// TwinCAT 3 PLC project CX7080_Robot_Controller
// ProgramVersion: 3.1.4024.0
// libraries:
//   Tc2_ModbusRTU, * (Beckhoff Automation GmbH)
//   Tc2_Standard, * (Beckhoff Automation GmbH)
//   Tc2_System, * (Beckhoff Automation GmbH)
//   Tc2_Utilities, * (Beckhoff Automation GmbH)
//   Tc3_Module, * (Beckhoff Automation GmbH)
// project tree:
//   DUTs/ eMbCycleState.TcDUT, eMbDiag.TcDUT, ST_HW_DI.TcDUT, ST_HW_DO.TcDUT, ST_MB_ReadRegs.TcDUT, ST_MB_WriteRegs.TcDUT, state_enum.TcDUT
//   GVLs/ GVL.TcGVL
//   / PlcTask.TcTTO
//   POUs/Comms/ FB_i_Watchdog.TcPOU, FB_ModbusComm.TcPOU, FB_Toggle_ReadWrite.TcPOU
//   POUs/ FB_Startup.TcPOU, I_JointJog.TcIO, MAIN.TcPOU, TESTING.TcPOU
//   POUs/Misc/ FB_System_Time.TcPOU
//   POUs/Motion/ FB_AutoSequence.TcPOU, FB_Jog_Joint.TcPOU, FB_Servo.TcPOU
//   POUs/Utilities/ FB_ElectromagnetActivate.TcPOU
// real-time tasks:
//   TASK PlcTask: cycle T#10ms, priority 20, ADS port 350
//   TASK PlcTask1: cycle T#10ms, priority 21, ADS port 351
//   TASK PlcTask2: cycle T#10ms, priority 22, ADS port 352
// I/O:
//   DEVICE Device 3 (CX7000), AmsNetId 5.140.122.236.4.1
//     Term 1 (CX7028) [CX7028-0000-0121]
//       modules: Module 1 (DIO_2x), Module 2 (Empty Module), Module 3 (DIO_2x), Module 4 (Empty Module), Module 5 (DI_2x), Module 6 (Empty Module), Module 7 (DI_2x), Module 8 (Empty Module)
//   DEVICE Device 1 (EtherCAT), AmsNetId 5.140.122.236.2.1
//     Term 1 (EK1200) [EK1200-7000 EtherCAT Power supply (1,5A E-Bus)]
//       Term 2 (EL1008) [EL1008 8Ch. Dig. Input 24V, 3ms]
//       Term 3 (EL1008) [EL1008 8Ch. Dig. Input 24V, 3ms]
//       Term 4 (EL2008) [EL2008 8Ch. Dig. Output 24V, 0.5A]
//       Term 5 (EL2008) [EL2008 8Ch. Dig. Output 24V, 0.5A]
//   DEVICE Device 7 (COM Port)
// variable links:
//   CX7080_Robot_Controller Instance <-> Device 1 (EtherCAT)/Term 1 (EK1200)/Term 2 (EL1008)
//     PlcTask Inputs/GVL.PB_EE_Grip <-> Channel 6/Input
//     PlcTask Inputs/GVL.PB_EE_Ungrip <-> Channel 8/Input
//     PlcTask Inputs/GVL.PB_J1_CCW <-> Channel 3/Input
//     PlcTask Inputs/GVL.PB_J2_CCW <-> Channel 5/Input
//     PlcTask Inputs/GVL.PB_J3_CCW <-> Channel 2/Input
//     PlcTask Inputs/GVL.PB_J1_CW <-> Channel 1/Input
//     PlcTask Inputs/GVL.PB_J2_CW <-> Channel 7/Input
//     PlcTask Inputs/GVL.PB_J3_CW <-> Channel 4/Input
//   CX7080_Robot_Controller Instance <-> Device 1 (EtherCAT)/Term 1 (EK1200)/Term 3 (EL1008)
//     PlcTask Inputs/GVL.PB_EMG_STOP <-> Channel 1/PB_EMG_STOP
//     PlcTask Inputs/GVL.PB_Record_Pos <-> Channel 3/PB_RECORD_POS
//     PlcTask Inputs/GVL.PB_Reset <-> Channel 2/PB_RESET
//     PlcTask Inputs/GVL.PB_Start_Pause <-> Channel 5/PB_START_PAUSE
//     PlcTask Inputs/GVL.SW_Jog_Auto <-> Channel 6/SW_JOG_AUTO
//     PlcTask Inputs/GVL.SW_Join_Cart <-> Channel 8/SW_JOINT_CART
//     PlcTask Inputs/GVL.SW_Slow_Fast <-> Channel 4/SW_SLOW_FAST
//   CX7080_Robot_Controller Instance <-> Device 1 (EtherCAT)/Term 1 (EK1200)/Term 4 (EL2008)
//     PlcTask Outputs/GVL.LED_EE_Grip <-> Channel 6/Output
//     PlcTask Outputs/GVL.LED_EE_Ungrip <-> Channel 8/Output
//     PlcTask Outputs/GVL.LED_J1_CCW <-> Channel 3/Output
//     PlcTask Outputs/GVL.LED_J2_CCW <-> Channel 5/Output
//     PlcTask Outputs/GVL.LED_J3_CCW <-> Channel 2/Output
//     PlcTask Outputs/GVL.LED_J1_CW <-> Channel 1/Output
//     PlcTask Outputs/GVL.LED_J2_CW <-> Channel 7/Output
//     PlcTask Outputs/GVL.LED_J3_CW <-> Channel 4/Output
//   CX7080_Robot_Controller Instance <-> Device 1 (EtherCAT)/Term 1 (EK1200)/Term 5 (EL2008)
//     PlcTask Outputs/GVL.LED_Comm_Fault <-> Channel 6/Output
//     PlcTask Outputs/GVL.LED_EMG_STOP <-> Channel 1/Output
//     PlcTask Outputs/GVL.LED_Record_Pos <-> Channel 3/Output
//     PlcTask Outputs/GVL.LED_Reset <-> Channel 2/Output
//     PlcTask Outputs/GVL.LED_Start_Pause <-> Channel 5/Output
//     PlcTask Outputs/GVL.LED_Warning <-> Channel 7/Output
//   CX7080_Robot_Controller Instance <-> Device 7 (COM Port)
//     PlcTask Inputs/MAIN.fb_ModbusComm.MB_Master.InData @bit {16..520 step 8} <-> Inputs/Data{1..64}  (64 links)
//     PlcTask Inputs/MAIN.fb_ModbusComm.MB_Master.InData <-> Inputs/Status
//     PlcTask Outputs/MAIN.fb_ModbusComm.MB_Master.OutData <-> Outputs/Ctrl
//     PlcTask Outputs/MAIN.fb_ModbusComm.MB_Master.OutData @bit {16..520 step 8} <-> Outputs/Data{1..64}  (64 links)

CONFIGURATION CX7080_Robot_Controller
    RESOURCE PLC ON TwinCAT3
        TASK PlcTask(INTERVAL := T#10ms, PRIORITY := 22);
        PROGRAM MAIN WITH PlcTask : MAIN;
    END_RESOURCE
END_CONFIGURATION

// ---- DUTs/eMbCycleState.TcDUT
{attribute 'namespace' := 'MyLib.Modbus'}
TYPE eMbCycleState :
(
    eMbState_Init,
    eMbState_Read,
    eMbState_Write,
    eMbState_Error
);
END_TYPE

// ---- DUTs/eMbDiag.TcDUT
TYPE eMbDiag :
(
    eMbDiag_Ok := 0,
    eMbDiag_Timeout := 1,
    eMbDiag_InvalidBusy := 2
);
END_TYPE

// ---- DUTs/ST_HW_DI.TcDUT
TYPE ST_HW_DI :
STRUCT
END_STRUCT
END_TYPE

// ---- DUTs/ST_HW_DO.TcDUT
TYPE ST_HW_DO :
STRUCT
END_STRUCT
END_TYPE

// ---- DUTs/ST_MB_ReadRegs.TcDUT
TYPE ST_MB_ReadRegs :
STRUCT
END_STRUCT
END_TYPE

// ---- DUTs/ST_MB_WriteRegs.TcDUT
TYPE ST_MB_WriteRegs :
STRUCT
END_STRUCT
END_TYPE

// ---- DUTs/state_enum.TcDUT
{attribute 'qualified_only'}
{attribute 'strict'}
TYPE state_enum :
(
	startup_mode,
	jog_joint_mode,
	jog_cartesian_mode,
	auto_mode,
	emg_stop_mode,
	comm_fault_mode,
	manual_mode
);
END_TYPE

// ---- GVLs/GVL.TcGVL
{attribute 'qualified_only'}
VAR_GLOBAL
	// Internal system parameters
	system_state : state_enum := state_enum.startup_mode; // Used to keep track of system state machine. Initialized in startup_mode.
	modbus_comm_fault : BOOL := FALSE;
	J1_Home_Pos : INT := 135; // Degrees
	J2_Home_Pos : INT := 135; // Degrees
	J3_Home_Pos : INT := 135; // Degrees
	LowSpeedSetting : REAL := 5; // [deg/s]
	HighSpeedSetting : REAL := 20; // [deg/s]
	
	BaseAngleMin : INT := 0;
	BaseAngleMax : INT := 180;
	ShoulderAngleMin : INT := 20;
	ShoulderAngleMax : INT := 120;
	ElbowAngleMin : INT := 0;
	ElbowAngleMax : INT := 180;
	
	// Inputs
	input1 AT %I* : BOOL;
	output1 AT %Q* : BOOL;
	PB_J1_CW AT %I* : BOOL;
	PB_J1_CCW AT %I*: BOOL;
	PB_J2_CW AT %I* : BOOL;
	PB_J2_CCW AT %I* : BOOL;
	PB_J3_CW AT %I* : BOOL;
	PB_J3_CCW AT %I* : BOOL;
	PB_EE_Grip AT %I* : BOOL;
	PB_EE_Ungrip AT %I* : BOOL;
	PB_EMG_STOP AT %I* : BOOL;
	PB_Reset AT %I* : BOOL;
	PB_Record_Pos AT %I* : BOOL;
	PB_Record_Delay AT %I* : BOOL;
	PB_Start_Pause AT %I* : BOOL;
	SW_Slow_Fast AT %I* : BOOL;
	SW_Join_Cart AT %I* : BOOL;
	SW_Jog_Auto AT %I* : BOOL;
	
	// Outputs
	LED_J1_CW AT %Q* : BOOL;
	LED_J1_CCW AT %Q*: BOOL;
	LED_J2_CW AT %Q* : BOOL;
	LED_J2_CCW AT %Q* : BOOL;
	LED_J3_CW AT %Q* : BOOL;
	LED_J3_CCW AT %Q* : BOOL;
	LED_EE_Grip AT %Q* : BOOL;
	LED_EE_Ungrip AT %Q* : BOOL;
	LED_EMG_STOP AT %Q* : BOOL;
	LED_Reset AT %Q* : BOOL;
	LED_Record_Pos AT %Q* : BOOL;
	LED_Record_Delay AT %Q* : BOOL;
	LED_Start_Pause AT %Q* : BOOL;
	LED_Comm_Fault AT %Q* : BOOL;
	LED_Warning AT %Q* : BOOL;
	
	// Modbus registers
	MB_Write_J1 : INT;
	MB_Write_J2 : INT;
	MB_Write_J3 : INT;
	MB_Write_Gripper : INT;
	MB_Write_Watchdog : INT;
	MB_Write_Blank1 : INT;
	MB_Write_Blank2 : INT;
	MB_Write_Blank3 : INT;
	MB_Write_Blank4 : INT;
	MB_Write_Blank5 : INT;
	MB_Read_Watchdog : INT;
	MB_Read_Blank2 : INT;
	MB_Read_Blank3 : INT;
	MB_Read_Blank4 : INT;
	MB_Read_Blank5 : INT;
	MB_Read_Blank6 : INT;
	MB_Read_Blank7 : INT;
	MB_Read_Blank8 : INT;
	MB_Read_Blank9 : INT;
	MB_Read_Blank10 : INT;
	
END_VAR

// ---- POUs/I_JointJog.TcIO
INTERFACE I_JointJog


(*
Hva er poenget med å bruke interface?
Det gjør separation of concerns enklere.
En funksjonsblokk trenger ikke å vite hvordan ting er implementert i (en annen funksjonsblokk?), men trenger
bare å kjenne til interface.
Dette gjør det enklere å drive med TDD (test driven development), da funksjonsblokker har mindre avhengigheter.


*)

METHOD Ramp : LREAL
VAR_INPUT
END_VAR
END_METHOD

END_INTERFACE

// ---- POUs/MAIN.TcPOU
PROGRAM MAIN
VAR
	fb_Startup : FB_Startup;
	fb_ModbusComm: FB_ModbusComm;
	fb_System_Time : FB_System_Time;
	fb_Jog_Joint : FB_Jog_Joint;
	fb_ElectromagnetActivate : FB_ElectromagnetActivate;
END_VAR


(*
GJENSTÅENDE ARBEID:
1) Implementer auto sekvens FB
2) 
*)


GVL.LED_J1_CW := GVL.PB_J1_CW;
GVL.LED_J2_CW := GVL.PB_J2_CW;
GVL.LED_J3_CW := GVL.PB_J3_CW;
GVL.LED_J1_CCW := GVL.PB_J1_CCW;
GVL.LED_J2_CCW := GVL.PB_J2_CCW;
GVL.LED_J3_CCW := GVL.PB_J3_CCW;
GVL.LED_EE_Grip := GVL.PB_EE_Grip;
GVL.LED_EE_Ungrip := GVL.PB_EE_Ungrip;
GVL.LED_EMG_STOP := NOT GVL.PB_EMG_STOP;
GVL.LED_Start_Pause := GVL.PB_Start_Pause;
GVL.LED_Reset := GVL.LED_Reset;
GVL.LED_Warning := TRUE;
GVL.LED_Reset := GVL.PB_Reset;
GVL.LED_Start_Pause := GVL.PB_Start_Pause;
GVL.LED_Record_Pos := GVL.PB_Record_Pos;


// Code which must run every PLC cycle.
fb_System_Time(); // Run FB to calculate Delta_Time


(* COMMENTING OUT FOR TESTING PURPOSES
IF NOT GVL.PB_EMG_STOP AND NOT (gvl.system_state = state_enum.startup_mode) THEN
	GVL.system_state := state_enum.emg_stop_mode;
ELSIF GVL.LED_Comm_Fault AND NOT (gvl.system_state = state_enum.startup_mode)  THEN
	GVL.system_state := state_enum.comm_fault_mode;
END_IF
*)


CASE gvl.system_state OF
state_enum.startup_mode:
	fb_Startup();
state_enum.jog_joint_mode:
	fb_Jog_Joint(
	lr_DeltaTime:= fb_ModbusComm.lreal_CycleTime, 
	lr_SlowModeVelocitySetting:= 1, 
	lr_FastModeVelovitySetting:= 10, 
	i_Base_LowLimit:= 0, 
	i_Base_HighLimit:= 180, 
	i_Shoulder_LowLimit:= 0, 
	i_Shoulder_HighLimit:= 180, 
	i_Elbow_LowLimit:= 0, 
	i_Elbow_HighLimit:= 180, 
	b_Enable_Servos:= TRUE, 
	SW_Fast_Mode:= GVL.SW_Slow_Fast, 
	PB_Base_Pos:= GVL.PB_J1_CCW, 
	PB_Base_Neg:= GVL.PB_J1_CW, 
	PB_Shoulder_Pos:= GVL.PB_J2_CCW, 
	PB_Shoulder_Neg:= GVL.PB_J2_CW, 
	PB_Elbow_Pos:= GVL.PB_J3_CCW, 
	PB_Elbow_Neg:= GVL.PB_J3_CW, 
	i_Set_Base=>, 
	i_Set_Shoulder=>, 
	i_Set_Elbow=>);
	
	fb_ElectromagnetActivate(
	b_activate := GVL.PB_EE_Grip,
	b_deactivate := GVL.PB_EE_Ungrip,
	b_CMD_Magnet =>);
	
state_enum.jog_cartesian_mode:
state_enum.manual_mode:
state_enum.emg_stop_mode:
state_enum.comm_fault_mode:
state_enum.auto_mode:
END_CASE

//fb_ModbusComm();
fb_ModbusComm(
	i_MBO_BaseAngle:= fb_Jog_Joint.i_Set_Base, 
	i_MBO_ShoulderAngle:= fb_Jog_Joint.i_Set_Shoulder, 
	i_MBO_ElbowAngle:= fb_Jog_Joint.i_Set_Elbow, 
	i_MBO_EndEffectorValue:= BOOL_TO_INT(fb_ElectromagnetActivate.b_CMD_Magnet), 
	b_MBO_EmergencyStop:= , 
	lreal_CycleTime := fb_System_Time.Delta_Time,
	iLastWrittenBaseAngle=> , 
	iLastWrittenShoulderAngle=> , 
	iLastWrittenElbowAngle=> , 
	b_MBI_LocalControl=> , 
	b_MBI_LocalEmergencyStopActive=> , 
	b_MBWatchdogTimeout=> GVL.LED_Comm_Fault, 
	i_MBI_LocalBaseAngle=> , 
	i_MBI_LocalShoulderAngle=> , 
	i_MBI_LocalElbowAngle=> , 
	i_MBI_LocalValueEndEffector=> );

END_PROGRAM

// ---- POUs/FB_Startup.TcPOU
FUNCTION_BLOCK FB_Startup
VAR_INPUT
END_VAR
VAR_OUTPUT
END_VAR
VAR
	timer1 : TON;
	timer2 : TON;
	timer3 : TON;
	timer4 : TON;
	timer5 : TON;
	timer6 : TON;
	timer7 : TON;
	EMG_STOP_RELEASED : BOOL;
END_VAR

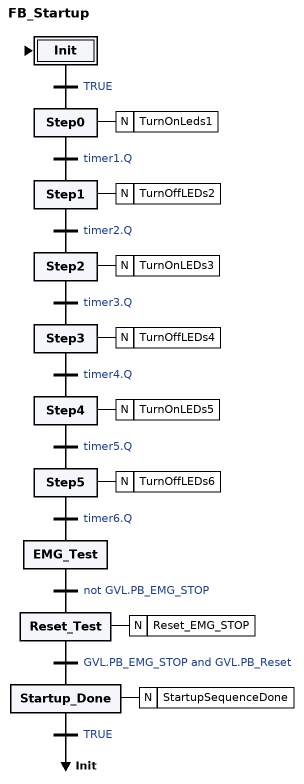
INITIAL_STEP Init:
END_STEP
TRANSITION FROM Init TO Step0
    := TRUE;
END_TRANSITION
STEP Step0:
    TurnOnLeds1(N);
END_STEP
TRANSITION FROM Step0 TO Step1
    := timer1.Q;
END_TRANSITION
STEP Step1:
    TurnOffLEDs2(N);
END_STEP
TRANSITION FROM Step1 TO Step2
    := timer2.Q;
END_TRANSITION
STEP Step2:
    TurnOnLEDs3(N);
END_STEP
TRANSITION FROM Step2 TO Step3
    := timer3.Q;
END_TRANSITION
STEP Step3:
    TurnOffLEDs4(N);
END_STEP
TRANSITION FROM Step3 TO Step4
    := timer4.Q;
END_TRANSITION
STEP Step4:
    TurnOnLEDs5(N);
END_STEP
TRANSITION FROM Step4 TO Step5
    := timer5.Q;
END_TRANSITION
STEP Step5:
    TurnOffLEDs6(N);
END_STEP
TRANSITION FROM Step5 TO EMG_Test
    := timer6.Q;
END_TRANSITION
STEP EMG_Test:
END_STEP
TRANSITION FROM EMG_Test TO Reset_Test
    := not GVL.PB_EMG_STOP;
END_TRANSITION
STEP Reset_Test:
    Reset_EMG_STOP(N);
END_STEP
TRANSITION FROM Reset_Test TO Startup_Done
    := GVL.PB_EMG_STOP and GVL.PB_Reset;
END_TRANSITION
STEP Startup_Done:
    StartupSequenceDone(N);
END_STEP
TRANSITION FROM Startup_Done TO Init
    := TRUE;
END_TRANSITION

METHOD AllLEDsTrigger : BOOL
VAR_INPUT
	OnOff : BOOL; // OnOff - Turn off, True - Turn On
END_VAR
GVL.LED_Comm_Fault := OnOff;
GVL.LED_EE_Grip := OnOff;
GVL.LED_EE_Ungrip := OnOff;
GVL.LED_EMG_STOP := OnOff;
GVL.LED_J1_CCW := OnOff;
GVL.LED_J1_CW := OnOff;
GVL.LED_J2_CCW := OnOff;
GVL.LED_J2_CW := OnOff;
GVL.LED_J3_CCW := OnOff;
GVL.LED_J3_CW := OnOff;
GVL.LED_Record_Delay := OnOff;
GVL.LED_Record_Pos := OnOff;
GVL.LED_Reset := OnOff;
GVL.LED_Start_Pause := OnOff;
GVL.LED_Warning := OnOff;
END_METHOD

ACTION Reset_EMG_STOP:
IF NOT GVL.PB_EMG_STOP THEN
	GVL.LED_EMG_STOP := TRUE;
END_IF

IF GVL.PB_EMG_STOP THEN
	GVL.LED_EMG_STOP := FALSE;
	GVL.LED_Reset := TRUE;
END_IF
END_ACTION

ACTION StartupSequenceDone:
GVL.LED_EMG_STOP := FALSE;
GVL.LED_Reset := FALSE;
GVL.system_state := state_enum.jog_joint_mode;
END_ACTION

ACTION TurnOffLEDs2:
timer1(IN := FALSE, PT := T#1S);
timer2(IN := TRUE, PT := T#1S);
timer3(IN := FALSE, PT := T#1S);
timer4(IN := FALSE, PT := T#1S);
timer5(IN := FALSE, PT := T#1S);
timer6(IN := FALSE, PT := T#1S);
timer7(IN := FALSE, PT := T#1S);
AllLEDsTrigger(FALSE);
END_ACTION

ACTION TurnOffLEDs4:
timer1(IN := FALSE, PT := T#1S);
timer2(IN := FALSE, PT := T#1S);
timer3(IN := FALSE, PT := T#1S);
timer4(IN := TRUE, PT := T#1S);
timer5(IN := FALSE, PT := T#1S);
timer6(IN := FALSE, PT := T#1S);
timer7(IN := FALSE, PT := T#1S);
AllLEDsTrigger(FALSE);
END_ACTION

ACTION TurnOffLEDs6:
timer1(IN := FALSE, PT := T#1S);
timer2(IN := FALSE, PT := T#1S);
timer3(IN := FALSE, PT := T#1S);
timer4(IN := FALSE, PT := T#1S);
timer5(IN := FALSE, PT := T#1S);
timer6(IN := TRUE, PT := T#1S);
timer7(IN := FALSE, PT := T#1S);
AllLEDsTrigger(FALSE);
END_ACTION

ACTION TurnOnLeds1:
timer1(IN := TRUE, PT := T#1S);
timer2(IN := FALSE, PT := T#1S);
timer3(IN := FALSE, PT := T#1S);
timer4(IN := FALSE, PT := T#1S);
timer5(IN := FALSE, PT := T#1S);
timer6(IN := FALSE, PT := T#1S);
timer7(IN := FALSE, PT := T#1S);
AllLEDsTrigger(TRUE);
END_ACTION

ACTION TurnOnLEDs3:
timer1(IN := FALSE, PT := T#1S);
timer2(IN := FALSE, PT := T#1S);
timer3(IN := TRUE, PT := T#1S);
timer4(IN := FALSE, PT := T#1S);
timer5(IN := FALSE, PT := T#1S);
timer6(IN := FALSE, PT := T#1S);
timer7(IN := FALSE, PT := T#1S);
AllLEDsTrigger(TRUE);
END_ACTION

ACTION TurnOnLEDs5:
timer1(IN := TRUE, PT := T#1S);
timer2(IN := FALSE, PT := T#1S);
timer3(IN := FALSE, PT := T#1S);
timer4(IN := FALSE, PT := T#1S);
timer5(IN := TRUE, PT := T#1S);
timer6(IN := FALSE, PT := T#1S);
timer7(IN := FALSE, PT := T#1S);
AllLEDsTrigger(TRUE);
END_ACTION

END_FUNCTION_BLOCK

// ---- POUs/Comms/FB_ModbusComm.TcPOU
FUNCTION_BLOCK FB_ModbusComm
VAR_INPUT
	i_MBO_BaseAngle : INT;
	i_MBO_ShoulderAngle : INT;
	i_MBO_ElbowAngle : INT;
	i_MBO_EndEffectorValue : INT;
	b_MBO_EmergencyStop : INT;
	lreal_CycleTime : LREAL;
END_VAR
VAR_OUTPUT
	iLastWrittenBaseAngle : INT;
	iLastWrittenShoulderAngle : INT;
	iLastWrittenElbowAngle : INT;
	b_MBI_LocalControl : BOOL;
	b_MBI_LocalEmergencyStopActive : BOOL;
	b_MBWatchdogTimeout : BOOL;
	i_MBI_LocalBaseAngle : INT;
	i_MBI_LocalShoulderAngle : INT;
	i_MBI_LocalElbowAngle : INT;
	i_MBI_LocalValueEndEffector : INT;
END_VAR
VAR
	i_MBO_WatchdogKick : INT;
	i_MBI_WatchdogBark : INT;
	MB_Master: ModbusRtuMaster_PcCOM;
	MB_ID: BYTE := 1;
	Data_Read : ARRAY[0..9] OF INT;
	Enable_Read: BOOL;
	Busy_Read: BOOL;
	Error_Read : BOOL;
	ErrorId_Read: Tc2_ModbusRTU.MODBUS_ERRORS;
	Register_Read_Address: WORD := 0;
	Data_Write : ARRAY[0..9] OF INT;
	Enable_Write: BOOL;
	Busy_Write: BOOL;
	Error_Write : BOOL;
	ErrorId_Write: Tc2_ModbusRTU.MODBUS_ERRORS;
	Register_Write_Address: WORD := 10;
	state : BOOL;
	Toggle_Auto : BOOL := TRUE;
	timer: TON;              // Timer On Delay function block
    clockSignal: BOOL := FALSE; // Output signal that toggles
    period: TIME := T#25MS;  // Period of the clock signal (1/10Hz = 100ms, so T#50ms for half-cycle)
	fb_i_Watchdog: FB_i_Watchdog;
	fb_Toggle_ReadWrite : FB_Toggle_ReadWrite;
END_VAR

fb_Toggle_ReadWrite(
	b_Enable_Write:= TRUE, 
	b_BusyRead:= Busy_Read, 
	b_BusyWrite:= Busy_Write, 
	b_Read=> Enable_Read, 
	b_Write=> Enable_Write);



MB_Master.ReadRegs(
    UnitID:= MB_ID, 
    Quantity:= 10, 
    MBAddr:= Register_Read_Address, 
    cbLength:= SIZEOF(Data_Read), 
    pMemoryAddr:= ADR(Data_Read), 
    Execute:= Enable_Read, 
    Timeout:= T#50MS, 
    BUSY=> Busy_Read, 
	
    Error=> Error_Read, 
    ErrorId=> ErrorId_Read, 
    cbRead=>);

	
	
i_MBI_LocalBaseAngle := Data_Read[0];
i_MBI_LocalShoulderAngle := Data_Read[1];
i_MBI_LocalBaseAngle := Data_Read[2];
i_MBI_LocalValueEndEffector := Data_Read[3];
b_MBI_LocalControl := INT_TO_BOOL(Data_Read[4]);
b_MBI_LocalEmergencyStopActive := INT_TO_BOOL(Data_Read[5]);
i_MBI_WatchdogBark := Data_Read[6];



Data_Write[0] := i_MBO_BaseAngle;
Data_Write[1] := i_MBO_ShoulderAngle;
Data_Write[2] := i_MBO_ElbowAngle;
Data_Write[3] := i_MBO_EndEffectorValue;
Data_Write[4] := b_MBO_EmergencyStop;
Data_Write[5] := i_MBO_WatchdogKick;


MB_Master.WriteRegs(
    UnitID:= MB_ID, 
    Quantity:= 10, 
    MBAddr:= Register_Write_Address, 
    cbLength:= SIZEOF(Data_Write), 
    pMemoryAddr:= ADR(Data_Write), 
    Execute:= Enable_Write, 
    Timeout:= T#50ms, 
    BUSY=> Busy_Write, 
    Error=> Error_Write, 
    ErrorId=> ErrorId_Write, 
    cbRead=>);



// Watchdog logic
i_MBO_WatchdogKick := i_MBO_WatchdogKick + 1;
IF i_MBO_WatchdogKick >= 1000 THEN
	i_MBO_WatchdogKick := 0;
END_IF

fb_i_Watchdog(
	lreal_MaxAllowedLatency:= 0.5, 
	i_Signal:= i_MBI_WatchdogBark, 
	lreal_dt:= lreal_CycleTime, 
	b_Timeout=> b_MBWatchdogTimeout, 
	lreal_AverageLatency=> );

END_FUNCTION_BLOCK

// ---- POUs/Comms/FB_i_Watchdog.TcPOU
FUNCTION_BLOCK FB_i_Watchdog
VAR_INPUT
	lreal_MaxAllowedLatency : LREAL; // [s]
	i_Signal : INT;
	lreal_dt : LREAL;
END_VAR
VAR_OUTPUT
	b_Timeout : BOOL;
	lreal_AverageLatency : LREAL; // Implement
END_VAR
VAR
	i_LastValue : INT;
	lreal_CurrentLatency : LREAL;
END_VAR

IF i_Signal <> i_LastValue THEN
	b_Timeout := FALSE;
	lreal_CurrentLatency := 0;
ELSE
	lreal_CurrentLatency := lreal_CurrentLatency + lreal_dt;
	IF lreal_CurrentLatency >= lreal_MaxAllowedLatency THEN
		b_Timeout := TRUE;
	END_IF
END_IF

i_LastValue := i_Signal;

END_FUNCTION_BLOCK

// ---- POUs/Comms/FB_Toggle_ReadWrite.TcPOU
FUNCTION_BLOCK FB_Toggle_ReadWrite
VAR_INPUT
	b_Enable_Write : BOOL;
	b_BusyRead : BOOL;
	b_BusyWrite : BOOL;
END_VAR
VAR_OUTPUT
	b_Read : BOOL;
	b_Write : BOOL;
END_VAR
VAR
	i_step : INT := 1; // Initially set to step 1
	F_TRIG_BusyRead : F_TRIG;
	F_TRIG_BusyWrite : F_TRIG;
END_VAR

F_TRIG_BusyRead(CLK:= b_BusyRead, Q=> );
F_TRIG_BusyWrite(CLK:= b_BusyWrite, Q=> );

CASE i_step OF
    1:
        b_Read := TRUE;
        b_Write := FALSE;
        i_step := 2;
    2:
        IF b_BusyRead THEN
            i_step := 3;
        END_IF
    3:
        b_Read := FALSE;
        i_step := 4;
    4:
        IF F_TRIG_BusyRead.Q THEN
            i_step := 5;
        END_IF
    5:
        IF b_Enable_Write THEN
            i_step := 7;
        ELSE
            i_step := 6;
        END_IF
    6:
        b_Read := TRUE;
        i_step := 2;
    7:
        b_Write := TRUE;
        b_Read := FALSE;
        i_step := 8;
    8:
        IF b_BusyWrite THEN
            i_step := 9;
        END_IF
    9:
        b_Write := FALSE;
        i_step := 10;
    10:
        IF F_TRIG_BusyWrite.Q THEN
            i_step := 1;
        END_IF
ELSE
    i_step := 1;
END_CASE

END_FUNCTION_BLOCK

// ---- POUs/Misc/FB_System_Time.TcPOU
FUNCTION_BLOCK FB_System_Time
VAR_OUTPUT
    Delta_Time : LREAL := 0;
	now : ULINT := 0;
END_VAR
VAR
    Last_Time : ULINT := 0;
	ConversionFactorSeconds : LREAL := 1E-7;
END_VAR

// FB must be called every PLC cycle, prefferably in the main() function.

now := Tc2_System.F_GetSystemTime();

IF Last_Time > 0 THEN
    Delta_Time := TO_LREAL(now - Last_Time) * ConversionFactorSeconds;
ELSE
    Delta_Time := 0;
END_IF

Last_Time := now;

END_FUNCTION_BLOCK

// ---- POUs/Motion/FB_Jog_Joint.TcPOU
FUNCTION_BLOCK FB_Jog_Joint
VAR_INPUT
	// Misc:
	lr_DeltaTime : LREAL;
	
	// Config parameters
	lr_SlowModeVelocitySetting : LREAL; // [deg/s]
	lr_FastModeVelovitySetting : LREAL; // [deg/s]
	i_Base_LowLimit : INT;
	i_Base_HighLimit : INT;
	i_Shoulder_LowLimit : INT;
	i_Shoulder_HighLimit : INT;
	i_Elbow_LowLimit : INT;
	i_Elbow_HighLimit : INT;
	
	
	
	// Control inputs
	b_Enable_Servos : BOOL;
	SW_Fast_Mode : BOOL; // True = fast mode, False = slow mode
	PB_Base_Pos : BOOL;
	PB_Base_Neg : BOOL;
	PB_Shoulder_Pos : BOOL;
	PB_Shoulder_Neg : BOOL;
	PB_Elbow_Pos : BOOL;
	PB_Elbow_Neg : BOOL;


END_VAR
VAR_OUTPUT
	i_Set_Base : INT;
	i_Set_Shoulder : INT;
	i_Set_Elbow : INT;
END_VAR
VAR
	lr_CurrentSpeedSetting : LREAL; // [deg/s]
	lr_Set_Base : LREAL;
	lr_Set_Shoulder : LREAL;
	lr_Set_Elbow : LREAL;
	
		// Structures:
	fb_Servo_Base : FB_Servo;
	fb_Servo_Shoulder : FB_Servo;
	fb_Servo_Elbow : FB_Servo;
END_VAR

fb_Servo_Base(
	b_EnableServo:= b_Enable_Servos, 
	b_CW:= PB_Base_Neg, 
	b_CCW:= PB_Base_Pos, 
	lr_deltaTime:= lr_DeltaTime, 
	lr_DegLowLim:= i_Base_LowLimit, 
	lr_DegHighLim:= i_Base_HighLimit, 
	lr_SlowModeVelocitySetting:= lr_SlowModeVelocitySetting, 
	lr_FastModeVelovitySetting:= lr_FastModeVelovitySetting, 
	SW_Fast_Mode:= SW_Fast_Mode, 
	i_Set_Angle=> i_Set_Base);

fb_Servo_Elbow(
	b_EnableServo:= b_Enable_Servos, 
	b_CW:= PB_Shoulder_Pos, 
	b_CCW:= PB_Shoulder_Neg, 
	lr_deltaTime:= lr_DeltaTime, 
	lr_DegLowLim:= i_Shoulder_LowLimit, 
	lr_DegHighLim:= i_Shoulder_HighLimit, 
	lr_SlowModeVelocitySetting:= lr_SlowModeVelocitySetting, 
	lr_FastModeVelovitySetting:= lr_FastModeVelovitySetting, 
	SW_Fast_Mode:= SW_Fast_Mode, 
	i_Set_Angle=> i_Set_Shoulder);

fb_Servo_Shoulder(
	b_EnableServo:= b_Enable_Servos, 
	b_CW:= PB_Elbow_Pos, 
	b_CCW:= PB_Elbow_Neg, 
	lr_deltaTime:= lr_DeltaTime, 
	lr_DegLowLim:= i_Elbow_LowLimit, 
	lr_DegHighLim:= i_Elbow_HighLimit, 
	lr_SlowModeVelocitySetting:= lr_SlowModeVelocitySetting, 
	lr_FastModeVelovitySetting:= lr_FastModeVelovitySetting, 
	SW_Fast_Mode:= SW_Fast_Mode, 
	i_Set_Angle=> i_Set_Elbow);

END_FUNCTION_BLOCK

// ---- POUs/Motion/FB_Servo.TcPOU
FUNCTION_BLOCK FB_Servo
VAR_INPUT
	b_EnableServo : BOOL;
	b_CW : BOOL;
	b_CCW : BOOL;
	lr_deltaTime : LREAL;
	lr_DegLowLim : INT;
	lr_DegHighLim : INT;
	lr_SlowModeVelocitySetting : LREAL; // [deg/s]
	lr_FastModeVelovitySetting : LREAL; // [deg/s]
	SW_Fast_Mode : BOOL; // True = fast mode, False = slow mode
END_VAR
VAR_OUTPUT
	i_Set_Angle : INT;
END_VAR
VAR
	lr_CurrentSpeedSetting : LREAL; // [deg/s]
	lr_Set_Angle : LREAL;
END_VAR

IF SW_Fast_Mode THEN
	lr_CurrentSpeedSetting := lr_FastModeVelovitySetting;
ELSE
	lr_CurrentSpeedSetting := lr_SlowModeVelocitySetting;
END_IF


IF b_EnableServo THEN
	IF b_CW AND NOT b_CCW THEN
		lr_Set_Angle := lr_Set_Angle + (lr_CurrentSpeedSetting * lr_deltaTime);
	ELSIF NOT b_CW AND b_CCW THEN
			lr_Set_Angle := lr_Set_Angle - (lr_CurrentSpeedSetting * lr_deltaTime);
	END_IF
	IF	lr_Set_Angle > lr_DegHighLim THEN
		lr_Set_Angle := lr_DegHighLim;
	ELSIF lr_Set_Angle < lr_DegLowLim THEN
		lr_Set_Angle := lr_DegLowLim;
	END_IF
	i_Set_Angle := LREAL_TO_INT(lr_Set_Angle);
END_IF;

END_FUNCTION_BLOCK

// ---- POUs/Utilities/FB_ElectromagnetActivate.TcPOU
FUNCTION_BLOCK FB_ElectromagnetActivate
VAR_INPUT
	b_activate : BOOL;
	b_deactivate : BOOL;
END_VAR
VAR_OUTPUT
	b_CMD_Magnet : BOOL;
END_VAR
VAR
END_VAR

(*
Spec:
Operator must hold activation button for a set amount of time before it changes from demagnectized to magnetized
Operator mudt hold deactivation button for a set amoint of time before it changes state from magnetized to demagnetized
If both magnetize button and demagnetize buttins are pressed simultanousely, nothing happens



TODO:
Implement debounce for buttons
Implement override release function to release magnetization on demand (for emergency situations)
*)

IF b_activate AND b_deactivate THEN
	// Do nothing - Operator should not push two buttons at the same time
ELSIF b_activate THEN
	b_CMD_Magnet := TRUE;
ELSIF b_deactivate THEN
	b_CMD_Magnet := FALSE;
END_IF

END_FUNCTION_BLOCK

// ---- POUs/Motion/FB_AutoSequence.TcPOU
FUNCTION_BLOCK FB_AutoSequence
VAR_INPUT
END_VAR
VAR_OUTPUT
END_VAR
VAR
END_VAR

(*
TODO
-Et punkt lagres ved å trykke på PB_RECORD_POS
-For å starte/pause en sekvens må PB_START_PAUSE trykkes inn
-Minst ett punkt må være lagret for å kunne starte en sekvens
-Hastighet kan enten være sakte eller rask, basert på bolsk verdi (false = slow, true = fast)
-For å slette lagrede mellombunkter, press og hold reset i tre sekunder
-Når sekvens er resatt, skal alle knapper blinke en gang





*)

END_FUNCTION_BLOCK

// ---- POUs/TESTING.TcPOU
PROGRAM TESTING
VAR
	Test_FB_Toggle_ReadWrite : FB_Toggle_ReadWrite;
END_VAR

Test_FB_Toggle_ReadWrite(
	b_Enable_Write:= , 
	b_BusyRead:= , 
	b_BusyWrite:= , 
	b_Read=> , 
	b_Write=> );

END_PROGRAM
